// TIA Portal V20 export
// export: Created 2026-10-20T18:55:49.0136215Z, ExportSetting None, DisplayName Totally Integrated Automation Portal, DisplayVersion V20 Update 6, DisplayName TIA Portal Openness, DisplayVersion V20 Update 6, DisplayName TIA Portal Version Control Interface, DisplayVersion V20 Update 6, DisplayName SINAMICS Startdrive Advanced, DisplayVersion V20 SP1, DisplayName SINAMICS Startdrive G130, G150, S120, S150, SINAMICS MV, G220, S200, S210, DisplayVersion V20 SP1, DisplayName SINAMICS Startdrive G110M, G120, G120C, G120D, G120P, G115D, DisplayVersion V20 SP1, DisplayName STEP 7 Professional, DisplayVersion V20 Update 6, DisplayName STEP 7 Safety, DisplayVersion V20 Update 2, DisplayName WinCC Basic/Comfort/Advanced, DisplayVersion V20 Update 6, DisplayName WinCC Unified, DisplayVersion V20 Update 6
VAR_GLOBAL   // PLC tag table "Lock_5"
   Lock_5_Estop_CH1 AT %I1790.2 : Bool;
   Lock_5_Closed_CH2 AT %I1790.1 : Bool;
   "Solenoid Enable_5" AT %Q1369.0 : Bool;
   Switches_5 AT %IB1277 : Byte;
   Lock_5_Estop_CH2 AT %I1790.3 : Bool;
   Lock_5_Closed_CH1 AT %I1790.0 : Bool;
   Lamps_5 AT %QB1363 : Byte;
   "Lock Reset_5" AT %Q1370.0 : Bool;
   Lock_5_Reset_Input2 AT %Q1791.1 : Bool;
   Lock_5_Reset_Input4 AT %Q1791.3 : Bool;
   Lock_5_Reset_Input3 AT %Q1791.2 : Bool;
   Lock_5_Reset_Input1 AT %Q1791.0 : Bool;
   "Guard Position_5" AT %I1278.0 : Bool;
   "Lock Position_5" AT %I1279.0 : Bool;
END_VAR
